// TIA Portal V20 export
Screen "02_Header"  1366x65
  ScreenItem "Dummy_ClockPulse" at 550,6 size 32x24  Type=HmiIOField
  ScreenItem "Dummy_Coordination" at 590,6 size 32x24  Type=HmiIOField
  ScreenItem "Backgroud_PermanentArea" at 0,0 size 1366x64  Type=HmiRectangle
  ScreenItem "Button_Manual" at 274,1 size 90x60  Type=HmiButton
  ScreenItem "Button_ControlOnOff" at 1,1 size 90x60  Type=HmiButton
  ScreenItem "Button_Start" at 92,1 size 90x60  Type=HmiButton
  ScreenItem "Button_Automatic" at 183,1 size 90x60  Type=HmiButton
  ScreenItem "Button_GoTo_AlarmHistory" at 1589,314 size 100x30  Type=HmiButton
  ScreenItem "Button_Special" at 1185,1 size 90x60  Type=HmiButton
  ScreenItem "Linie_1" at 91,1 size 0x60  Type=HmiLine
  ScreenItem "Linie_2" at 182,1 size 0x60  Type=HmiLine
  ScreenItem "Linie_3" at 273,1 size 0x60  Type=HmiLine
  ScreenItem "Linie_Left" at 0,1 size 0x60  Type=HmiLine
  ScreenItem "Linie_Right" at 1275,1 size 0x60  Type=HmiLine
  ScreenItem "auto_Blocked" at 184,4 size 14x14  Type=HmiGraphicView
  ScreenItem "start_Foreground_Blocked" at 93,2 size 90x61  Type=HmiGraphicView
  ScreenItem "start_Blocked" at 93,4 size 14x14  Type=HmiGraphicView
  ScreenItem "auto_Foreground_Blocked" at 184,2 size 90x61  Type=HmiGraphicView
  ScreenItem "manual_Foreground_Blocked" at 275,1 size 90x62  Type=HmiGraphicView
  ScreenItem "manual_Blocked" at 275,4 size 14x14  Type=HmiGraphicView
  ScreenItem "Silence button" at 1005,1 size 90x60  Type=HmiButton
  ScreenItem "Fusszeile_Button_Nav1" at 1275,1 size 90x60  Type=HmiButton
  ScreenItem "Button_GoTo_AlarmHistory_1" at 1394,314 size 100x30  Type=HmiButton
  ScreenItem "Text_1" at 1394,103 size 75x28  Type=HmiText
  ScreenItem "DateTime" at 838,33 size 162x24  Type=HmiIOField
  ScreenItem "IOField_ProjectName" at 538,0 size 460x30  Type=HmiIOField
  ScreenItem "RF1060R_PMLOGON" at 594,35 size 34x22  Type=HmiFaceplateContainer
  ScreenItem "HMI_No" at 544,35 size 28x25  Type=HmiFaceplateContainer
  ScreenItem "SMC_Diag" at 574,35 size 18x21  Type=HmiFaceplateContainer
  ScreenItem "DeviceDiag_Summary" at 669,35 size 32x22  Type=HmiFaceplateContainer
  ScreenItem "PLC_Checksum" at 630,35 size 28x22  Type=HmiFaceplateContainer
  ScreenItem "Button_GoTo_SystemSettings" at 544,28 size 114x30  Type=HmiButton
  ScreenItem "Button_GoTo_DemoSlide" at 544,-4 size 461x30  Type=HmiButton
  ScreenItem "Button_OPModeSelect" at 365,3 size 173x59  Type=HmiButton
  ScreenItem "Button_GoTo_PN-Diag" at 667,30 size 36x30  Type=HmiButton
  ScreenItem "Linie_4" at 364,1 size 0x60  Type=HmiLine
  ScreenItem "Linie_5" at 539,1 size 0x60  Type=HmiLine
  ScreenItem "Opmode_24" at 365,0 size 173x63  Type=HmiFaceplateContainer
  ScreenItem "Faceplate container_1" at 703,26 size 100x35  Type=HmiFaceplateContainer
  ScreenItem "Button_GoTo_AlarmHistory_2" at 677,38 size 100x30  Type=HmiButton
  ScreenItem "Button_Ack_BackgroundAnimation" at 1094,1 size 90x60  Type=HmiButton
  ScreenItem "OPmodeArea_Selected" at 1120,38 size 38x24  Type=HmiFaceplateContainer
  ScreenItem "Linie_6" at 1093,1 size 0x60  Type=HmiLine
  ScreenItem "Linie_7" at 1184,1 size 0x60  Type=HmiLine
  ScreenItem "Button_Ack" at 1095,2 size 90x60  Type=HmiButton
